Staubli VAL3: utBorder.dtx

public string sBorderColour
